(*
SPDX-FileCopyrightText: © 2026 Oleksandr Tiutyk <trofimich@gmail.com>
SPDX-License-Identifier: MIT
License: https://opensource.org/license/mit
*)

(*!
<summary>
Beckhoff EL3356: 1-channel precise resistor bridge / load cell terminal (24-bit).
</summary>
<description>
Requires the one-channel strain-gauge INT32 assignment: status PDO 0x1A00, value PDO 0x1A01,
and control PDO 0x1600. Keep both input PDOs enabled and link Status and Value separately.
Value is signed calculated load; engineering scaling follows calibration. REAL load, two-channel voltage,
optional filter-frequency and timestamp PDOs are outside this model; disable or link optional PDOs separately.
When used for I/O, link located fields or their containing buffers to the matching selected PDOs.
The record is not a packed wire buffer; compiler padding is not part of the device specification.
Unlinked/default values do not prove valid I/O. The caller evaluates bus/channel validity before use.
Use one owner task per instance and externally synchronize other access; multi-field snapshots are not atomic.
Copies store data without creating hardware links. Keep borrowed field references valid while consumers are bound.
This passive record performs no validation, synchronization, configuration or protocol advancement.
</description>
*)
TYPE EL3356 :
STRUCT
	Ch1 : STRAIN_GAUGE_CHANNEL;
END_STRUCT
END_TYPE

(* stored: Version 1.1.0.1, ProductVersion 3.1.4026.20
   DUT EL3356: Id {2bef32b3-f1e0-4555-8d21-ed39d697c8d9} *)
